Fanuc KAREL source: KO00011.KL

PROGRAM KO00011
%NOLOCKGROUP
VAR
  P1: XYZWPR
  P2: XYZWPR
  P3: XYZWPR
  OUT: XYZWPREXT
BEGIN
  OUT = FRAME(P1, P2, P3)
END KO00011
